Staubli VAL3: getIndex.pgx

public program getIndex(string x_sKey, num& x_nIndex)
  local bool l_bResult
  local num l_nIndex
begin
  toNum(x_sKey,l_nIndex,l_bResult)
  if l_bResult
    x_nIndex=l_nIndex
  else
    x_nIndex=-1
    userPageAlert("未选择有效项目！")
  endIf
end
